// TIA Portal V19 export
DATA_BLOCK "VFD_1"   // DB84
// stored: InstanceOfName VFD_DATA, InstanceOfType FB
"VFD_DATA"
   // VAR_INPUT
   //    ON_OFF : Bool;
   //    RESET : Bool;
   //    SPEED_SP : Real;
   // END_VAR
   // VAR_OUTPUT
   //    READY : Bool;
   //    RUNNING : Bool;
   //    TRIP : Bool;
   //    ACT_SPEED : Real;
   //    "LOCAL/REMOTE" : Int;
   // END_VAR
   // VAR_IN_OUT
   //    DATA : "VFD";
   // END_VAR
BEGIN
END_DATA_BLOCK
